Fanuc KAREL source: kx00015.KL

-- PROVISIONAL review KL for V770-1; original PC SHA256 cd4d95bdebc15dcade8c36f1187960f48235148ecaf5c3dab7b69571a51e5597
-- Incomplete behavior may be omitted. Consult companion uncertainty JSON. Do not deploy.
PROGRAM KX00015
%NOLOCKGROUP
VAR
  I : INTEGER
  J : INTEGER
  B : BOOLEAN
  F : FILE
  S : STRING[80]
-- UNRESOLVED_DECL P type=000102
BEGIN
  -- UNRESOLVED_PC offsets 5-7; opcodes 9D,0E
  -- UNRESOLVED_PC offsets 12-16; opcodes 7F
END KX00015
